Staubli VAL3: simulateTRAJ.pgx

program simulateTRAJ(string x_sKey)
begin
  call simulate:simulateTRAJ(x_sKey)
end
